(* IEC 61131-3 sources: plc-repo-template/src/POUs/FB_Example, 2 files *)

(* ---- FB_Example.decl.st ---- *)
// Назначение: пример ФБ устройства — двухпозиционный регулятор с гистерезисом
//             (насос подкачки по уровню): включение при значении не выше
//             (уставка - гистерезис), отключение при значении не ниже уставки.
//             Режимы E_DeviceMode, безопасное состояние (выход отключён) при отказе
//             измерения, квитирование отказа, счётчик включений для оценки износа.
// Автор:      kr0nsch
// Версия:     0.1.0
// Документ:   docs/ARCHITECTURE.md, раздел «Пример в src/»
FUNCTION_BLOCK FB_Example IMPLEMENTS I_Resettable
VAR_INPUT
    // режим работы; пока режим не назначен — выведено из работы
    eMode : E_DeviceMode := E_DeviceMode.OutOfService;
    rValue_pct : REAL;          // измеренное значение, % диапазона датчика
    xValueValid : BOOL;         // измерение достоверно (например, по NAMUR NE 43)
    rSetpoint_pct : REAL := GVL_Const.EXAMPLE_SP_DEFAULT_PCT;       // уставка отключения, %
    rHysteresis_pct : REAL := GVL_Const.EXAMPLE_HYST_DEFAULT_PCT;   // гистерезис ниже уставки, %
    xManualOn : BOOL;           // команда «включить» в ручном режиме
END_VAR
VAR_OUTPUT
    xOut : BOOL;                // TRUE — исполнительный механизм включён
    xFault : BOOL;              // отказ измерения зафиксирован, нужен вызов Acknowledge()
    rSetpointUsed_pct : REAL;   // уставка после ограничения диапазоном, %
    rHysteresisUsed_pct : REAL; // гистерезис после ограничения диапазоном, %
END_VAR
VAR
    xOutPrev : BOOL;            // выход в предыдущем вызове — для счёта включений по фронту
    udiCount : UDINT;           // число включений выхода с последнего Reset()
END_VAR

(* ---- FB_Example.impl.st ---- *)
// 1. Параметры оператора ограничиваем допустимыми диапазонами из GVL_Const
rSetpointUsed_pct := F_Clamp(rValue := rSetpoint_pct,
                             rLow := GVL_Const.EXAMPLE_SP_MIN_PCT,
                             rHigh := GVL_Const.EXAMPLE_SP_MAX_PCT);
rHysteresisUsed_pct := F_Clamp(rValue := rHysteresis_pct,
                               rLow := GVL_Const.EXAMPLE_HYST_MIN_PCT,
                               rHigh := GVL_Const.EXAMPLE_HYST_MAX_PCT);

// 2. Отказ измерения фиксируем в авторежиме — только там измерение управляет выходом.
//    Защёлка: отказ держится до квитирования, даже если измерение восстановилось.
xFault := xFault OR (eMode = E_DeviceMode.Auto AND NOT xValueValid);

// 3. Выход по режимам
CASE eMode OF
    E_DeviceMode.Auto:
        IF xFault THEN
            xOut := FALSE;      // безопасное состояние до квитирования
        ELSIF rValue_pct <= rSetpointUsed_pct - rHysteresisUsed_pct THEN
            xOut := TRUE;
        ELSIF rValue_pct >= rSetpointUsed_pct THEN
            xOut := FALSE;
        END_IF
        // внутри зоны гистерезиса выход сохраняет прежнее состояние

    E_DeviceMode.Manual:
        xOut := xManualOn;

    E_DeviceMode.Local, E_DeviceMode.OutOfService:
        // местный пост управляет сам, вывод из работы — команда ПЛК снимается
        xOut := FALSE;

ELSE
    xOut := FALSE;              // неизвестное значение режима — безопасное состояние
END_CASE

// 4. Счёт включений по переднему фронту выхода; на пределе счётчик не переполняется
IF xOut AND NOT xOutPrev AND udiCount < GVL_Const.EXAMPLE_COUNT_MAX THEN
    udiCount := udiCount + 1;
END_IF
xOutPrev := xOut;
